Fanuc KAREL source: NC0064.KL

PROGRAM NC0064
%NOLOCKGROUP
ROUTINE R
VAR
  X : INTEGER
  I1 : INTEGER
  I2 : INTEGER
  I3 : INTEGER
BEGIN
  X = 1
  FOR I1 = 1 TO 2 DO
    FOR I2 = 1 TO 2 DO
      FOR I3 = 1 TO 2 DO
        X = X + 1
      ENDFOR
    ENDFOR
  ENDFOR
END R
BEGIN
  R
END NC0064
